FUNCTION_BLOCK SCALE_CLAMP (* Migrated from IEC 61131-3 ST *)
  (* Standard: 61499-2 *)
  (* Version 1.0, 2026-11-06, st2fb *)
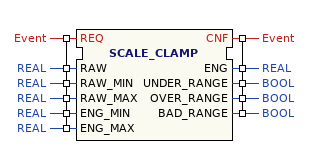
  EVENT_INPUT
    REQ WITH RAW, RAW_MIN, RAW_MAX, ENG_MIN, ENG_MAX;
  END_EVENT
  EVENT_OUTPUT
    CNF WITH ENG, UNDER_RANGE, OVER_RANGE, BAD_RANGE;
  END_EVENT
  VAR_INPUT
    RAW : REAL;
    RAW_MIN : REAL;
    RAW_MAX : REAL;
    ENG_MIN : REAL;
    ENG_MAX : REAL;
  END_VAR
  VAR_OUTPUT
    ENG : REAL;
    UNDER_RANGE : BOOL;
    OVER_RANGE : BOOL;
    BAD_RANGE : BOOL;
  END_VAR
  VAR
    SPAN : REAL;
  END_VAR
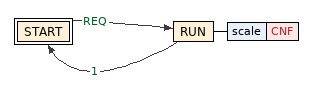
  EC_STATES
    START;
    RUN : scale -> CNF;
  END_STATES
  EC_TRANSITIONS
    START TO RUN := REQ;
    RUN TO START := 1;
  END_TRANSITIONS
  ALGORITHM scale IN ST:
SPAN := RAW_MAX - RAW_MIN;
BAD_RANGE := SPAN <= 0.0;
IF BAD_RANGE THEN
  ENG := ENG_MIN;
  UNDER_RANGE := FALSE;
  OVER_RANGE := FALSE;
ELSE
  UNDER_RANGE := RAW < RAW_MIN;
  OVER_RANGE := RAW > RAW_MAX;
  IF UNDER_RANGE THEN
    ENG := ENG_MIN;
  ELSIF OVER_RANGE THEN
    ENG := ENG_MAX;
  ELSE
    ENG := ENG_MIN + (RAW - RAW_MIN) * (ENG_MAX - ENG_MIN) / SPAN;
  END_IF;
END_IF;
  END_ALGORITHM
END_FUNCTION_BLOCK
